FUNCTION_BLOCK BasicAdapter2 (* Adapter communication, events only *)
  (* Standard: 61499-2; Description: Copyright (c) 2023 Johannes Kepler University Linz This program and the accompanying materials are made available under the terms of the Eclipse Public License 2.0 which is available at https://www.eclipse.org/legal/epl-2.0/ SPDX-License-Identifier: EPL-2.0 *)
  (* Version 1.0, 2023-03-07, Bianca Wiesmayr, Johannes Kepler University Linz, initial API and implementation and/or initial documentation *)
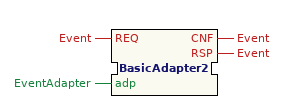
  EVENT_INPUT
    REQ;
  END_EVENT
  EVENT_OUTPUT
    CNF;
    RSP;
  END_EVENT
  SOCKETS
    adp : EventAdapter;
  END_SOCKETS
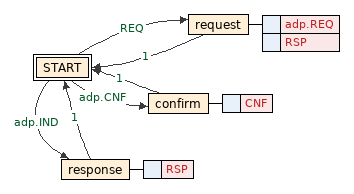
  EC_STATES
    START; (* Initial State *)
    request : -> adp.REQ, -> RSP;
    confirm : -> CNF;
    response : -> RSP;
  END_STATES
  EC_TRANSITIONS
    START TO request := REQ;
    request TO START := 1;
    START TO confirm := adp.CNF;
    START TO response := adp.IND;
    response TO START := 1;
    confirm TO START := 1;
  END_TRANSITIONS
END_FUNCTION_BLOCK
